NAMESPACE TiaMcp_UnitA
DATA_BLOCK "TgpUnit_GlobalTimer"
{ S7_Optimized_Access := 'TRUE' }
VERSION : 0.1
"IEC_TIMER"
BEGIN
END_DATA_BLOCK
END_NAMESPACE
